VISUALIZATION Header  // 1024x768
END_VISUALIZATION

(* stored: Version 1.1.0.1
   Visu Header: Id {ff4a00ff-3a67-4255-86ce-c2cd9274ddf2} *)
